Yaskawa INFORM job: CONFPRO.JBI

/JOB
//NAME CONFPRO
//POS
///NPOS 8,0,0,0,0,0
///TOOL 9
///POSTYPE PULSE
///PULSE
C00000=0,-19456,25243,0,27307,0
C00001=333592,-19456,25243,202752,27307,-151924
C00002=-333592,-116736,126216,-202752,-27307,208193
C00003=18032,38912,-37865,42685,-45511,33761
C00004=-306544,87552,-56797,-181410,81920,-100720
C00005=-306544,87552,-56797,-181410,81920,-100720
C00006=333592,-19456,25243,202752,27307,-151924
C00007=-333592,-116736,126216,-202752,-27307,208193
//INST
<volatile>
///COMM Generated using RoboDK
///ATTR SC,RW
///GROUP1 RB1
NOP
'Program generated by RoboDK v
'6.0.7 for Yaskawa Motoman DX1
'350D on XX/XX/XXXX 18:00:00
'Using nominal kinematics.
'Using Frame S (targets wrt ba
'se):
'1234.6,-98.8,50.5,0.0,0.0,30.
'0
'Tool Tool S should be close t
'o:
'10.0,20.0,150.0,0.0,0.0,0.0
MOVL C00000 V=100.0
MOVL C00001 V=100.0
MOVL C00002 V=100.0
MOVJ C00003 VJ=50.00
MOVJ C00004 VJ=50.00
MOVC C00005 V=100.0
MOVC C00006 V=100.0
MOVC C00007 V=100.0
END
